(* IEC 61131-3 sources: kns-port-domestic/upstream/kns-pump-station/src/POUs/Log/F_UtcNowMs, 2 files *)

(* ---- F_UtcNowMs.decl.st ---- *)
// Назначение: текущее время UTC, мс от 1970 (SysTimeRtcHighResGet) для меток журнала и списка тревог;
//             0 — часы недоступны или не выставлены (время раньше LOG_UTC_MIN_MS).
// Автор:      kr0nsch
// Версия:     0.1.0
// Документ:   docs/DESIGN.md, разделы 9.1, 9.3
FUNCTION F_UtcNowMs : ULINT
VAR
    uliNow_ms : ULINT;              // ответ часов реального времени
END_VAR

(* ---- F_UtcNowMs.impl.st ---- *)
IF SysTimeRtcHighResGet(pTimestamp := uliNow_ms) = GVL_Const.LOG_RTC_OK
   AND uliNow_ms >= GVL_Const.LOG_UTC_MIN_MS THEN
    F_UtcNowMs := uliNow_ms;
ELSE
    F_UtcNowMs := 0;
END_IF
